(* IEC 61131-3 sources: model-first-plc-agent-ai/results/T2-W-27, 2 files *)

(* ---- a1_code.st ---- *)
FUNCTION_BLOCK FillingRuntime
VAR_INPUT
    start : BOOL;
    stop : BOOL;
    LSH : BOOL;
    LSHH : BOOL;
    TimerDuration : TIME;
END_VAR
VAR_OUTPUT
    fill_valve : BOOL;
    discharge_valve : BOOL;
END_VAR
VAR
    x0 : BOOL := TRUE;
    x1 : BOOL := FALSE;
    timer_done : BOOL := FALSE;
    FillingTimer : TON;
END_VAR

(* Transition t1: enter the filling step. *)
IF x0 AND start AND NOT stop AND NOT LSHH THEN
    x0 := FALSE;
    x1 := TRUE;
END_IF;

(* The timer measures the activity of x1, including its entry scan. *)
FillingTimer(IN := x1, PT := TimerDuration);
timer_done := FillingTimer.Q;

(* Transition t2: return to the initial step. *)
IF x1 AND (stop OR LSHH OR timer_done) THEN
    x1 := FALSE;
    x0 := TRUE;

    (* Reset the owned timer when its step becomes inactive. *)
    FillingTimer(IN := FALSE, PT := TimerDuration);
    timer_done := FALSE;
END_IF;

fill_valve := x1;
discharge_valve := FALSE;

END_FUNCTION_BLOCK

PROGRAM Main
VAR
    StartCommand AT %IX100.0 : BOOL;
    StopCommand AT %IX100.1 : BOOL;
    LSH AT %IX100.2 : BOOL;
    LSHH AT %IX100.3 : BOOL;
    FillValve AT %QX100.0 : BOOL;
    DischargeValve AT %QX100.1 : BOOL;
END_VAR
VAR
    (* Configurable filling-duration parameter. *)
    TimerDuration : TIME := T#5s;
    StartEdge : R_TRIG;
    FillingControl : FillingRuntime;
END_VAR

StartEdge(CLK := StartCommand);

FillingControl(
    start := StartEdge.Q,
    stop := StopCommand,
    LSH := LSH,
    LSHH := LSHH,
    TimerDuration := TimerDuration
);

FillValve := FillingControl.fill_valve;
DischargeValve := FillingControl.discharge_valve;

END_PROGRAM

(* ---- a2_code.st ---- *)
FUNCTION_BLOCK FB_TimedTankFilling
VAR_INPUT
    StartCommand : BOOL;
    StopCommand : BOOL;
    LSH : BOOL;
    LSHH : BOOL;
    TimerDuration : TIME;
END_VAR
VAR_OUTPUT
    fill_valve : BOOL;
    discharge_valve : BOOL;
END_VAR
VAR
    StartEdge : R_TRIG;
    FillingTimer : TON;
    ActiveState : INT := 0;
    start : BOOL := FALSE;
    stop : BOOL := FALSE;
    timer_done : BOOL := FALSE;
END_VAR

StartEdge(CLK := StartCommand);
start := StartEdge.Q;
stop := StopCommand;

IF stop THEN
    ActiveState := 0;
ELSE
    CASE ActiveState OF
        0:
            IF start THEN
                ActiveState := 1;
            END_IF;
        1:
            ActiveState := 1;
    ELSE
        ActiveState := 0;
    END_CASE;
END_IF;

FillingTimer(
    IN := (ActiveState = 1),
    PT := TimerDuration
);
timer_done := FillingTimer.Q;

IF ActiveState = 1 THEN
    IF stop OR timer_done OR LSHH THEN
        ActiveState := 0;
        FillingTimer(IN := FALSE, PT := TimerDuration);
        timer_done := FillingTimer.Q;
    END_IF;
END_IF;

fill_valve := (ActiveState = 1);
discharge_valve := FALSE;

END_FUNCTION_BLOCK

PROGRAM Main
VAR
    StartCommand AT %IX100.0 : BOOL;
    StopCommand AT %IX100.1 : BOOL;
    LSH AT %IX100.2 : BOOL;
    LSHH AT %IX100.3 : BOOL;
    FillValve AT %QX100.0 : BOOL;
    DischargeValve AT %QX100.1 : BOOL;
END_VAR
VAR
    TankController : FB_TimedTankFilling;
    TimerDuration : TIME := T#10s;
END_VAR

TankController(
    StartCommand := StartCommand,
    StopCommand := StopCommand,
    LSH := LSH,
    LSHH := LSHH,
    TimerDuration := TimerDuration
);

FillValve := TankController.fill_valve;
DischargeValve := TankController.discharge_valve;

END_PROGRAM
